(* IEC 61131-3 sources: plc-vscode/tests/st/all/trust-platform/conformance/cases/memory_map/cfm_memory_map_wildcard_unresolved_002, 1 file *)

(* ---- program.st ---- *)
PROGRAM Main
VAR
    out AT %M* : BOOL;
END_VAR

out := TRUE;
END_PROGRAM
